Fanuc KAREL source: kd00025.KL

-- PROVISIONAL review KL for V1013-1; original PC SHA256 96e8bde2ade2769e310bae85db5beae533bc6aa480d1f241389852f486a3feda
-- Incomplete behavior may be omitted. Consult companion uncertainty JSON. Do not deploy.
PROGRAM KD00025
%NOLOCKGROUP
VAR
  I : INTEGER
  J : INTEGER
  B : BOOLEAN
  R : REAL
  S : STRING[80]
BEGIN
  -- UNRESOLVED_PC offsets 5-31; opcodes 9D,2E,25,81,18,9D,1B,9D,12,22,9D,13,04
  -- UNRESOLVED_PC offsets 36-40; opcodes 7F
END KD00025
